// TIA Portal V20 export
// export: Created 2026-10-20T18:55:45.054484Z, ExportSetting None, DisplayName Totally Integrated Automation Portal, DisplayVersion V20 Update 6, DisplayName TIA Portal Openness, DisplayVersion V20 Update 6, DisplayName TIA Portal Version Control Interface, DisplayVersion V20 Update 6, DisplayName SINAMICS Startdrive Advanced, DisplayVersion V20 SP1, DisplayName SINAMICS Startdrive G130, G150, S120, S150, SINAMICS MV, G220, S200, S210, DisplayVersion V20 SP1, DisplayName SINAMICS Startdrive G110M, G120, G120C, G120D, G120P, G115D, DisplayVersion V20 SP1, DisplayName STEP 7 Professional, DisplayVersion V20 Update 6, DisplayName STEP 7 Safety, DisplayVersion V20 Update 2, DisplayName WinCC Basic/Comfort/Advanced, DisplayVersion V20 Update 6, DisplayName WinCC Unified, DisplayVersion V20 Update 6
VAR_GLOBAL   // PLC tag table "Lock_3"
   Lock_3_Estop_CH1 AT %I1774.2 : Bool;
   Lock_3_Closed_CH1 AT %I1774.0 : Bool;
   Switches_3 AT %IB902 : Byte;
   Lamps_3 AT %QB1066 : Byte;
   "Lock Reset_3" AT %Q1073.0 : Bool;
   Lock_3_Estop_CH2 AT %I1774.3 : Bool;
   Lock_3_Closed_CH2 AT %I1774.1 : Bool;
   "Solenoid Enable_3" AT %Q1072.0 : Bool;
   Lock_3_Reset_Input3 AT %Q1775.2 : Bool;
   Lock_3_Reset_Input1 AT %Q1775.0 : Bool;
   Lock_3_Reset_Input4 AT %Q1775.3 : Bool;
   Lock_3_Reset_Input2 AT %Q1775.1 : Bool;
   "Lock Position_3" AT %I1163.0 : Bool;
   "Guard Position_3" AT %I903.0 : Bool;
END_VAR
